// Résultat d'une commande (docs/05 § 2, docs/06 § 6.1)
{attribute 'qualified_only'}
{attribute 'strict'}
TYPE E_CmdResult :
(
    None := 0,
    Accepted := 1,
    Rejected := 2
) USINT;
END_TYPE

(* stored: Version 1.1.0.1, ProductVersion 3.1.4024.12
   DUT E_CmdResult: Id {e4a32a2e-1de6-54a6-b3c0-2dc009c0f4f1} *)
